Fanuc KAREL source: ka00092.KL

-- PROVISIONAL review KL for V940-1; original PC SHA256 06e199ae2f2235b782ef07e0babb58691ff2f27b2fdb7ca8013935cc0d30d2dc
-- Incomplete behavior may be omitted. Consult companion uncertainty JSON. Do not deploy.
PROGRAM KA00092
%NOLOCKGROUP
-- UNRESOLVED_DECL SRC type=000199
-- UNRESOLVED_DECL DST type=000199
BEGIN
  -- V9_ZERO_TABLE_METADATA_HINT layout=0001; no indexed target words; source/name/runtime held
  -- UNRESOLVED_PC offsets 5-20; opcodes 49,4A
  -- UNRESOLVED_PC offsets 25-29; opcodes 7F
END KA00092
